{attribute 'qualified_only'}
VAR_GLOBAL
	// Robot Position for Unity (0-100)
    MyRobotY : REAL ;
END_VAR

(* stored: Version 1.1.0.1, ProductVersion 3.1.4024.15
   GVL GVL_GamePong: Id {2a8087ec-579f-4382-bca8-837c68c9ea88} *)
